(* IEC 61131-3 sources: llm-plc-st-eval/data/definitivo/qwen2.5-coder_14b/C8/zero_shot, 3 files *)

(* ---- ejec_1.st ---- *)
```pascal
FUNCTION_BLOCK FB_Valvula
VAR_INPUT
    nivelAlto : BOOL; // Entrada que indica el nivel alto
END_VAR

VAR_OUTPUT
    valvula : BOOL; // Salida que controla la válvula
END_VAR

VAR
    T1 : TON; // Temporizador de retardo por encendido
END_VAR

// Inicialización del temporizador T1 con un tiempo preestablecido de 5 segundos
IF nivelAlto THEN
    T1(IN := nivelAlto, PT := T#5S);
END_IF;

// La válvula se activa cuando el temporizador T1 ha terminado
valvula := T1.Q;
```

Este código en Structured Text (ST) implementa el comportamiento descrito en el Ladder Diagram. La variable `nivelAlto` es la entrada que indica el nivel alto, y `valvula` es la salida que controla la válvula. El temporizador `T1` se configura con un tiempo preestablecido de 5 segundos (`T#5S`). La válvula se activa cuando el temporizador `T1` ha terminado su cuenta.

(* ---- ejec_2.st ---- *)
```pascal
FUNCTION_BLOCK FB_Valvula
VAR_INPUT
    nivelAlto : BOOL; // Entrada que indica el nivel alto
END_VAR

VAR_OUTPUT
    valvula : BOOL; // Salida que controla la válvula
END_VAR

VAR
    T1 : TON; // Temporizador de tipo TON
END_VAR

// Inicialización del temporizador T1 con un tiempo preestablecido de 5 segundos
T1.PT := T#5S;

// Rama 1: Si nivelAlto es verdadero, arranca el temporizador T1
IF nivelAlto THEN
    T1(IN := TRUE);
ELSE
    T1(IN := FALSE);
END_IF;

// Rama 2: Si el temporizador T1 ha terminado, activa la válvula
valvula := T1.Q;
```

Este código en Structured Text (ST) implementa el comportamiento descrito en el Ladder Diagram, utilizando un temporizador de tipo TON (Timer On Delay) para controlar la válvula. La variable `nivelAlto` es la entrada que indica el nivel alto, y `valvula` es la salida que controla la válvula. El temporizador `T1` se configura con un tiempo preestablecido de 5 segundos.

(* ---- ejec_3.st ---- *)
```pascal
FUNCTION_BLOCK FB_Valvula
VAR_INPUT
    nivelAlto : BOOL; // Entrada que indica el nivel alto
END_VAR

VAR_OUTPUT
    valvula : BOOL; // Salida que controla la válvula
END_VAR

VAR
    T1 : TON; // Temporizador de retardo por encendido
END_VAR

// Inicialización del temporizador T1 con un tiempo preestablecido de 5 segundos
IF nivelAlto THEN
    T1(IN := TRUE, PT := T#5S);
ELSE
    T1(IN := FALSE);
END_IF;

// La válvula se abre cuando el temporizador T1 ha terminado su cuenta
valvula := T1.Q;
```

Este código en Structured Text (ST) implementa el comportamiento descrito en el Ladder Diagram, utilizando un temporizador de retardo por encendido (TON) para controlar la válvula. La variable `nivelAlto` es la entrada que indica el nivel alto, y `valvula` es la salida que controla la válvula. El temporizador `T1` tiene un tiempo preestablecido de 5 segundos.
